Fanuc KAREL source: KA00204.KL

PROGRAM KA00204
%NOLOCKGROUP
VAR
  SRC: ARRAY[4] OF VECTOR
  DST: ARRAY[4] OF SHORT
BEGIN
  DST = SRC
END KA00204
